(*
SPDX-FileCopyrightText: © 2026 Oleksandr Tiutyk <trofimich@gmail.com>
SPDX-License-Identifier: MIT
License: https://opensource.org/license/mit
*)

(*!
<summary>
Beckhoff SSI absolute encoder channel process image.
</summary>
<description>
Represents the SSI 32-bit position and two-byte status variant.
EL5001 requires firmware 11 or later and selection of the two-byte status PDO (0x1A01).
Earlier EL5001 firmware supports only one status byte and is incompatible with this channel.
For EL5002 select the corresponding two-byte status PDO for each channel. No byte-status conversion occurs.
When used for I/O, link located fields or their containing buffers to the matching selected PDOs.
The record is not a packed wire buffer; compiler padding is not part of the device specification.
Unlinked/default values do not prove valid I/O. The caller evaluates bus/channel validity before use.
Use one owner task per instance and externally synchronize other access; multi-field snapshots are not atomic.
Copies store data without creating hardware links. Keep borrowed field references valid while consumers are bound.
This passive record performs no validation, synchronization, configuration or protocol advancement.
</description>
*)
TYPE SSI_ENCODER_CHANNEL :
STRUCT
	Status AT %I* : WORD;
	Value AT %I* : UDINT;
END_STRUCT
END_TYPE

(* stored: Version 1.1.0.1, ProductVersion 3.1.4026.20
   DUT SSI_ENCODER_CHANNEL: Id {91fa5d19-9c3b-4370-9de9-d68aea8f1cc9} *)
